(* IEC 61131-3 sources: other-plc-idf/examples/open_linux/counter, 1 file *)

(* ---- main.st ---- *)
(* Real IEC ST example. No physical I/O or network access. *)
PROGRAM MAIN
VAR
    COUNTER : DINT := 0;
    HEARTBEAT : BOOL := FALSE;
END_VAR
COUNTER := COUNTER + 1;
IF (COUNTER MOD 10) = 0 THEN
    HEARTBEAT := NOT HEARTBEAT;
END_IF;
END_PROGRAM

CONFIGURATION Config0
RESOURCE Res0 ON PLC
    TASK scan (INTERVAL := T#20ms, PRIORITY := 0);
    PROGRAM instance0 WITH scan : MAIN;
END_RESOURCE
END_CONFIGURATION
